TYPE ST_FireflyToUnity :
STRUCT
    fX : REAL;   // -100..+100 %, 0 = home (middle of the scene), +100 = right edge of the garden
    fY : REAL;   // -100..+100 %, 0 = home (middle of the scene), +100 = top edge (robot forward)
END_STRUCT
END_TYPE

(* stored: Version 1.1.0.1, ProductVersion 3.1.4024.15
   DUT ST_FireflyToUnity: Id {9d301b2d-3137-4776-92dc-e9c35f7115e9} *)
